// TIA Portal V20 export
// export: Created 2026-10-19T18:36:57.7500855Z, ExportSetting WithDefaults, DisplayName Totally Integrated Automation Portal, DisplayVersion V20 Update 6, DisplayName TIA Portal Openness, DisplayVersion V20 Update 6, DisplayName TIA Portal Version Control Interface, DisplayVersion V20 Update 6, DisplayName SINAMICS Startdrive Advanced, DisplayVersion V20 SP1, DisplayName SINAMICS Startdrive G130, G150, S120, S150, SINAMICS MV, G220, S200, S210, DisplayVersion V20 SP1, DisplayName SINAMICS Startdrive G110M, G120, G120C, G120D, G120P, G115D, DisplayVersion V20 SP1, DisplayName STEP 7 Professional, DisplayVersion V20 Update 6, DisplayName STEP 7 Safety, DisplayVersion V20 Update 2, DisplayName WinCC Basic/Comfort/Advanced, DisplayVersion V20 Update 6, DisplayName WinCC Unified, DisplayVersion V20 Update 6
DATA_BLOCK "Conveyor_HMI_FB_1_DB"   // DB15
VERSION : 0.1
// stored: AutoNumber true, DBAccessibleFromOPCUA true, InstanceOfName Conveyor_HMI_FB_1, InstanceOfType FB
"Conveyor_HMI_FB_1"
   // VAR_INPUT
   //    HMI_No : UInt;
   //    Sys_No : UInt;
   //    Zone : UInt;
   // END_VAR
   // VAR_IN_OUT
   //    Enable : Bool;
   //    Mode_Change : UInt;
   //    Transfer_To_ID : DInt;
   //    Transfer_From_ID : DInt;
   //    "Enable(1)" : Bool;
   //    "Mode_Change(1)" : UInt;
   //    "Transfer_To_ID(1)" : DInt;
   //    "Transfer_From_ID(1)" : DInt;
   // END_VAR
   // VAR
   //    R_Charge_Cnv_Commands { S7_SetPoint := 'True'} : R_TRIG;
   //    T_Reset_Charge { S7_SetPoint := 'True'} : TON_TIME;
   //    ID { S7_SetPoint := 'True'} : DInt;
   //    "ID(1)" : DInt;
   //    ID_Old { S7_SetPoint := 'True'} : DInt;
   //    "ID_Old(1)" : DInt;
   // END_VAR
BEGIN
END_DATA_BLOCK
